FUNCTION "Feed_BCNV_Cnv2(1)_1"   // FC 30, author

VAR_INPUT
   HMI_No : UInt;
   System_No : UInt;
   Level : UInt;
   Light_Guard_IO : Bool;
END_VAR

VAR_OUTPUT
   Light_Guard_Bypass : Bool;
END_VAR

   // RETURN : Void
BEGIN
//Sensors
"CNV_HMI"."Left(1)"[#HMI_No] := "Control_DB".LCnv_Sys[#System_No].Cnv_Level[#Level].Cnv2.Inputs.Left;
"CNV_HMI"."Lpd1(1)"[#HMI_No] := "Control_DB".LCnv_Sys[#System_No].Cnv_Level[#Level].Cnv2.Inputs.Lpd1;
"CNV_HMI"."Lpd2(1)"[#HMI_No] := "Control_DB".LCnv_Sys[#System_No].Cnv_Level[#Level].Cnv2.Inputs.Lpd2;
"CNV_HMI"."Right(1)"[#HMI_No] := "Control_DB".LCnv_Sys[#System_No].Cnv_Level[#Level].Cnv2.Inputs.Right;
"CNV_HMI"."Rpd1(1)"[#HMI_No] := "Control_DB".LCnv_Sys[#System_No].Cnv_Level[#Level].Cnv2.Inputs.Rpd1;
"CNV_HMI"."Rpd2(1)"[#HMI_No] := "Control_DB".LCnv_Sys[#System_No].Cnv_Level[#Level].Cnv2.Inputs.Rpd2;
"CNV_HMI"."Sdetect1(1)"[#HMI_No] := "Control_DB".LCnv_Sys[#System_No].Cnv_Level[#Level].Cnv2.Inputs.Sdetect1;
"CNV_HMI"."Sdetect2(1)"[#HMI_No] := "Control_DB".LCnv_Sys[#System_No].Cnv_Level[#Level].Cnv2.Inputs.Sdetect2;
"HMI_Light_Guard" := #Level = 1; //To show the button
IF "Control_DB".LCnv_Sys[#System_No].Cnv_Level[#Level].Cnv2.Safety_Stop_Cnrl.Inputs.DP_Extended AND
    NOT "Control_DB".LCnv_Sys[#System_No].Cnv_Level[#Level].Cnv2.Safety_Stop_Cnrl.Inputs.DP_Retracted THEN
    "CNV_HMI"."UpDown(1)"[#HMI_No] := 1;
ELSIF NOT "Control_DB".LCnv_Sys[#System_No].Cnv_Level[#Level].Cnv2.Safety_Stop_Cnrl.Inputs.DP_Extended AND
    "Control_DB".LCnv_Sys[#System_No].Cnv_Level[#Level].Cnv2.Safety_Stop_Cnrl.Inputs.DP_Retracted THEN
    "CNV_HMI"."UpDown(1)"[#HMI_No] := 2;
ELSE
    "CNV_HMI"."UpDown(1)"[#HMI_No] := 0;
END_IF;

//Status
"CNV_HMI"."Mode(1)"[#HMI_No] := "Control_DB".LCnv_Sys[#System_No].Cnv_Level[#Level].Cnv2.Mode;
"CNV_HMI"."Enabled(1)"[#HMI_No] := "Control_DB".LCnv_Sys[#System_No].Cnv_Level[#Level].Cnv2.Enabled;
"CNV_HMI"."Error(1)"[#HMI_No] := "Control_DB".LCnv_Sys[#System_No].Cnv_Level[#Level].Cnv2.Error;
"CNV_HMI"."Warning(1)"[#HMI_No] := "Control_DB".LCnv_Sys[#System_No].Cnv_Level[#Level].Cnv2.Warning;
"CNV_HMI"."Stopped(1)"[#HMI_No] := "Control_DB".LCnv_Sys[#System_No].Cnv_Level[#Level].Cnv2.Stopped;
"CNV_HMI"."Running(1)"[#HMI_No] := "Control_DB".LCnv_Sys[#System_No].Cnv_Level[#Level].Cnv2.Running;
"CNV_HMI"."Ready_For_Task(1)"[#HMI_No] := "Control_DB".LCnv_Sys[#System_No].Cnv_Level[#Level].Cnv2.Ready_For_Task;
"CNV_HMI"."Occupied(1)"[#HMI_No] := "Control_DB".LCnv_Sys[#System_No].Cnv_Level[#Level].Cnv2.Cnv_Occupied;
"CNV_HMI"."Shuttle_in_place(1)"[#HMI_No] := "Control_DB".LCnv_Sys[#System_No].Cnv_Level[#Level].Cnv2.Shuttle_In_Place;
"CNV_HMI"."Current_Task_Type(1)"[#HMI_No] := "Control_DB".LCnv_Sys[#System_No].Cnv_Level[#Level].Cnv2.Current_Task_Type;
"CNV_HMI"."Task_ID(1)"[#HMI_No] := "Control_DB".LCnv_Sys[#System_No].Cnv_Level[#Level].Cnv2.Current_Task_ID;
"CNV_HMI"."SM_State(1)"[#HMI_No] := "Control_DB".LCnv_Sys[#System_No].Cnv_Level[#Level].Cnv2.SM_State;
"CNV_HMI"."Pallet_Type(1)"[#HMI_No] := "Control_DB".LCnv_Sys[#System_No].Cnv_Level[#Level].Cnv2.Pallet_Type;
IF "Control_DB".LCnv_Sys[#System_No].Cnv_Level[#Level].Cnv2.Motor.Forward THEN
    "CNV_HMI"."Motor_Direction(1)"[#HMI_No] := 1;
ELSIF "Control_DB".LCnv_Sys[#System_No].Cnv_Level[#Level].Cnv2.Motor.Reverse THEN
    "CNV_HMI"."Motor_Direction(1)"[#HMI_No] := 2;
ELSE
    "CNV_HMI"."Motor_Direction(1)"[#HMI_No] := 0;
END_IF;
"CNV_HMI"."Motor_Speed_Requested(1)"[#HMI_No] := "Control_DB".LCnv_Sys[#System_No].Cnv_Level[#Level].Cnv2.Motor.Speed;
"CNV_HMI"."Motor_Speed_Actual(1)"[#HMI_No] := "Control_DB".LCnv_Sys[#System_No].Cnv_Level[#Level].Cnv2.Motor.Speed_Actual;
"CNV_HMI"."Motor_Ready(1)"[#HMI_No] := "Control_DB".LCnv_Sys[#System_No].Cnv_Level[#Level].Cnv2.Motor.Ready;
"CNV_HMI"."Motor_Current_Actual(1)"[#HMI_No] := "Control_DB".LCnv_Sys[#System_No].Cnv_Level[#Level].Cnv2.Motor.Actual_Current;
"CNV_HMI"."Motor_Actual_Torque(1)"[#HMI_No] := "Control_DB".LCnv_Sys[#System_No].Cnv_Level[#Level].Cnv2.Motor.Actual_Torque;
"CNV_HMI"."Transfer_To_ID(1)"[#HMI_No] := "Control_DB".LCnv_Sys[#System_No].Cnv_Level[#Level].Cnv2.Instruction.Transfer_To_ID;
"CNV_HMI"."Transfer_From_ID(1)"[#HMI_No] := "Control_DB".LCnv_Sys[#System_No].Cnv_Level[#Level].Cnv2.Instruction.Transfer_From_ID;

IF "Control_DB".LCnv_Sys[#System_No].Cnv_Level[#Level].Cnv2.Motor.Error THEN
    "CNV_HMI"."Motor_Status(1)"[#HMI_No] := 2;
ELSIF "Control_DB".LCnv_Sys[#System_No].Cnv_Level[#Level].Cnv2.Motor.Enabled THEN
    "CNV_HMI"."Motor_Status(1)"[#HMI_No] := 1;
ELSIF NOT "Control_DB".LCnv_Sys[#System_No].Cnv_Level[#Level].Cnv2.Motor.Enabled THEN
    "CNV_HMI"."Motor_Status(1)"[#HMI_No] := 0;
END_IF;

//Instructions
"Control_DB".LCnv_Sys[#System_No].Cnv_Level[#Level].Cnv2.Instruction.Stop := "CNV_HMI"."Stop(1)"[#HMI_No];
"Control_DB".LCnv_Sys[#System_No].Cnv_Level[#Level].Cnv2.Instruction.Execute := "CNV_HMI"."Manual_Fwd(1)"[#HMI_No] OR "CNV_HMI"."Manual_Bwd(1)"[#HMI_No];
"Control_DB".LCnv_Sys[#System_No].Cnv_Level[#Level].Cnv2.Instruction.Mode_Change := "CNV_HMI"."Mode_Change(1)"[#HMI_No];
"Control_DB".LCnv_Sys[#System_No].Cnv_Level[#Level].Cnv2.Instruction.Enable := "CNV_HMI"."Enable(1)"[#HMI_No];
#Light_Guard_Bypass := "HMI_Light_Guard_Bypass";

"Control_DB".LCnv_Sys[#System_No].Cnv_Level[#Level].Cnv2.Instruction.Reset := "CNV_HMI"."Reset(1)"[#HMI_No] OR "Screen_DB_1".Reset_All[#HMI_No];
IF "Control_DB".LCnv_Sys[#System_No].Cnv_Level[#Level].Cnv2.Mode <> 3 THEN
    "Control_DB".LCnv_Sys[#System_No].Cnv_Level[#Level].Cnv2.Instruction.Foward := "CNV_HMI"."Manual_Fwd(1)"[#HMI_No];
    "Control_DB".LCnv_Sys[#System_No].Cnv_Level[#Level].Cnv2.Instruction.Backward := "CNV_HMI"."Manual_Bwd(1)"[#HMI_No];
    "Control_DB".LCnv_Sys[#System_No].Cnv_Level[#Level].Cnv2.Instruction.Start_Transfer := "CNV_HMI"."Start_Transfer(1)"[#HMI_No];
    "Control_DB".LCnv_Sys[#System_No].Cnv_Level[#Level].Cnv2.Safety_Stop_Cnrl.Instruction.Manual_Extend := "CNV_HMI"."Manual_Sfty_Stopper_Up(1)"[#HMI_No];
    "Control_DB".LCnv_Sys[#System_No].Cnv_Level[#Level].Cnv2.Safety_Stop_Cnrl.Instruction.Manual_Retract := "CNV_HMI"."Manual_Sfty_Stopper_Down(1)"[#HMI_No];
    "Control_DB".LCnv_Sys[#System_No].Cnv_Level[#Level].Cnv2.Instruction.Task_ID := "CNV_HMI"."Task_ID(1)"[#HMI_No];
    "Control_DB".LCnv_Sys[#System_No].Cnv_Level[#Level].Cnv2.Instruction.Pallet_Align_Left := "CNV_HMI"."Pallet_Align_Left(1)"[#HMI_No];
    "Control_DB".LCnv_Sys[#System_No].Cnv_Level[#Level].Cnv2.Instruction.Pallet_Align_Right := "CNV_HMI"."Pallet_Align_Right(1)"[#HMI_No];
    IF "CNV_HMI"."Mode_Change(1)"[#HMI_No] <> 2 THEN
        "Control_DB".LCnv_Sys[#System_No].Cnv_Level[#Level].Cnv2.Instruction.Pallet_Allignment := "CNV_HMI"."Pallet_Allignment(1)"[#HMI_No] := FALSE;
    ELSE
        "Control_DB".LCnv_Sys[#System_No].Cnv_Level[#Level].Cnv2.Instruction.Pallet_Allignment := "CNV_HMI"."Pallet_Allignment(1)"[#HMI_No];
    END_IF;
    IF "CNV_HMI".In_Out[#System_No] THEN // 0 = ECNV RECEIVE, 1 = ECONV SEND
        "Control_DB".LCnv_Sys[#System_No].Cnv_Level[#Level].Cnv2.Instruction.Transfer_To_ID := 0;
        "Control_DB".LCnv_Sys[#System_No].Cnv_Level[#Level].Cnv2.Instruction.Transfer_From_ID := DINT#120000 + (#Level * 100) + #System_No;
    ELSE
        "Control_DB".LCnv_Sys[#System_No].Cnv_Level[#Level].Cnv2.Instruction.Transfer_To_ID := DINT#120000 + (#Level * 100) + #System_No;
        "Control_DB".LCnv_Sys[#System_No].Cnv_Level[#Level].Cnv2.Instruction.Transfer_From_ID := 0;
    END_IF;
END_IF;

END_FUNCTION